// TIA Portal V21 program export: 0 tag tables, 0 data types, 0 data blocks, 2 code blocks (in call order from the OBs), 0 instance data blocks

ORGANIZATION_BLOCK "Pair"   // OB1, LAD
BEGIN

REGION Network 1: Motor
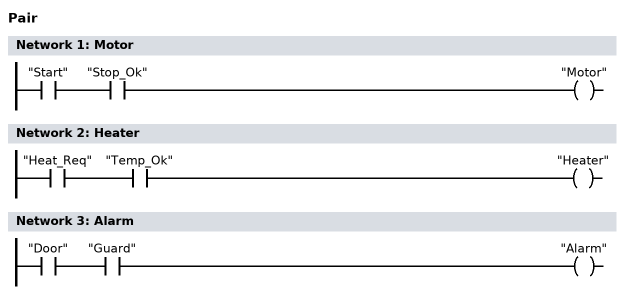
   RUNG wire#powerrail
      Contact( "Start" )
      Contact( "Stop_Ok" )
      Coil( "Motor" )
   END_RUNG
   // the same network as SCL:
   "Motor" := "Start" AND "Stop_Ok";
END_REGION

REGION Network 2: Heater
   RUNG wire#powerrail
      Contact( "Heat_Req" )
      Contact( "Temp_Ok" )
      Coil( "Heater" )
   END_RUNG
   // the same network as SCL:
   "Heater" := "Heat_Req" AND "Temp_Ok";
END_REGION

REGION Network 3: Alarm
   RUNG wire#powerrail
      Contact( "Door" )
      Contact( "Guard" )
      Coil( "Alarm" )
   END_RUNG
   // the same network as SCL:
   "Alarm" := "Door" AND "Guard";
END_REGION
END_ORGANIZATION_BLOCK

FUNCTION_BLOCK "Mixed"   // FB1, LAD
BEGIN

REGION Network 1: Unknown part
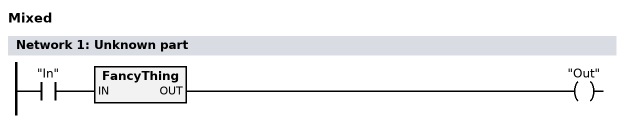
   // no SCL statement known for FancyThing: written as a call
   "Out" := FancyThing("In");
END_REGION

REGION Network 2 (SCL): SCL inside
END_REGION

REGION Network 3: Empty
END_REGION
END_FUNCTION_BLOCK
